// Maps a severity onto a TMC event (event class + event id).
INTERFACE I_EventEntryProvider

METHOD GetEventEntry : TcEventEntry
VAR_INPUT
	eSeverity	: TcEventSeverity;
END_VAR
END_METHOD

END_INTERFACE

(* stored: Version 1.1.0.1, ProductVersion 3.1.4026.26
   Itf I_EventEntryProvider: Id {7e757470-ce7b-413d-8f35-d886c49b9f56}
   Method GetEventEntry: Id {c70d9519-63eb-4c3c-bad5-e30305ce9996} *)
